// TIA Portal V20 export
FUNCTION_BLOCK "POS3_0_Antriebe"   // FB34, FBD
{ S7_Optimized_Access := 'TRUE' }
// stored: MemoryReserve 100, SetENOAutomatically false
   VAR
      "-1001T1_OM_PRM_Access_Instance" { S7_SetPoint := 'True'} : "OM_PRM_Access";
      "-1001T1_Oriental" { S7_SetPoint := 'True'} : "Oriental_AZD-KPN_Profinet";
      "-1002T2_OM_PRM_Access_Instance" { S7_SetPoint := 'True'} : "OM_PRM_Access";
      "-1002T2_Oriental_Drehachse" { S7_SetPoint := 'True'} : "Oriental_AZD-KPN_Profinet";
      Pos_Alt { S7_SetPoint := 'True'} : Real;
      Delta : Real;
   END_VAR
BEGIN

REGION Network 1 (SCL): -1001T1 Pos 3.0 Positionierachse Vorgaben Geschwindigkeit und Beschleunigung
   "POS3_0_Signal"."-1001T1 Oriental_Beschleunigung" := 50.0;
   "POS3_0_Signal"."-1001T1 Oriental_Speed" := 100.0;
END_REGION

REGION Network 2 (SCL): -1001T1 Pos 3.0 Positionierachse Achse stopp
   // Achse stopp
   IF "03_Betriebsart_DB"."Schutztüren OK" AND
       "DE_POS3_0_Endlage_Überlastzylinder" THEN
       "POS3_0_Signal"."-1001T1 Oriental_Steuerung".E_STOP := FALSE;
   ELSE
       "POS3_0_Signal"."-1001T1 Oriental_Steuerung".E_STOP := TRUE;
   END_IF;
END_REGION

REGION Network 3 (SCL): -1001T1 Pos 3.0 Positionierachse Position 0 Achse [Grundstellung]
   "POS3_0_Signal"."-1001T1 Oriental_Positionen".Operation_type[0] := 16#0001;
   "POS3_0_Signal"."-1001T1 Oriental_Positionen".Soll_Position[0] := 0.0;
   "POS3_0_Signal"."-1001T1 Oriental_Positionen".Geschwindigkeit[0] := 10.0;
   "POS3_0_Signal"."-1001T1 Oriental_Positionen".Start_Rampe[0] := "POS3_0_Signal"."-1001T1 Oriental_Beschleunigung"; // Start-Rampe %
   "POS3_0_Signal"."-1001T1 Oriental_Positionen".Stopp_Rampe[0] := "POS3_0_Signal"."-1001T1 Oriental_Beschleunigung"; // Stopp-Rampe %
   "POS3_0_Signal"."-1001T1 Oriental_Positionen".Arbeitsstrom[0] := 100;  // Arbeitsstrom in %
   "POS3_0_Signal"."-1001T1 Oriental_Positionen".Positioniertoleranz[0] := 0.02;
END_REGION

REGION Network 4 (SCL): -1001T1 Pos 3.0 Positionierachse Position 1 Achse [GS aus Verwaltung]
   "POS3_0_Signal"."-1001T1 Oriental_Positionen".Operation_type[1] := 16#0001;

   "POS3_0_Signal"."-1001T1 Oriental_Positionen".Start_Rampe[1] := "POS3_0_Signal"."-1001T1 Oriental_Beschleunigung"; // Start-Rampe %
   "POS3_0_Signal"."-1001T1 Oriental_Positionen".Stopp_Rampe[1] := "POS3_0_Signal"."-1001T1 Oriental_Beschleunigung"; // Stopp-Rampe %
   "POS3_0_Signal"."-1001T1 Oriental_Positionen".Arbeitsstrom[1] := 100;   // Arbeitsstrom in %
   "POS3_0_Signal"."-1001T1 Oriental_Positionen".Positioniertoleranz[1] := 0.02;
END_REGION

REGION Network 5 (SCL): -1001T1 Pos 3.0 Positionierachse Position 2 Achse [AS aus Verwaltung]
   "POS3_0_Signal"."-1001T1 Oriental_Positionen".Operation_type[2] := 16#0001;

   "POS3_0_Signal"."-1001T1 Oriental_Positionen".Start_Rampe[2] := "POS3_0_Signal"."-1001T1 Oriental_Beschleunigung"; // Start-Rampe %
   "POS3_0_Signal"."-1001T1 Oriental_Positionen".Stopp_Rampe[2] := "POS3_0_Signal"."-1001T1 Oriental_Beschleunigung"; // Stopp-Rampe %
   "POS3_0_Signal"."-1001T1 Oriental_Positionen".Arbeitsstrom[2] := 100;  // Arbeitsstrom in %
   "POS3_0_Signal"."-1001T1 Oriental_Positionen".Positioniertoleranz[2] := 0.02;
END_REGION

REGION Network 6 (SCL): -1001T1 Pos 3.0 Positionierachse Position 3 Achse
   "POS3_0_Signal"."-1001T1 Oriental_Positionen".Operation_type[3] := 16#0001;

   "POS3_0_Signal"."-1001T1 Oriental_Positionen".Start_Rampe[3] := "POS3_0_Signal"."-1001T1 Oriental_Beschleunigung" ; // Start-Rampe %
   "POS3_0_Signal"."-1001T1 Oriental_Positionen".Stopp_Rampe[3] := "POS3_0_Signal"."-1001T1 Oriental_Beschleunigung" ; // Stopp-Rampe %
   "POS3_0_Signal"."-1001T1 Oriental_Positionen".Arbeitsstrom[3] := 100; // Arbeitsstrom in %
   "POS3_0_Signal"."-1001T1 Oriental_Positionen".Positioniertoleranz[3] := 0.02;
END_REGION

REGION Network 7 (SCL): -1001T1 Pos 3.0 Positionierachse Position 4 Achse
   "POS3_0_Signal"."-1001T1 Oriental_Positionen".Operation_type[4] := 16#0001;

   "POS3_0_Signal"."-1001T1 Oriental_Positionen".Start_Rampe[4] := "POS3_0_Signal"."-1001T1 Oriental_Beschleunigung" ; // Start-Rampe %
   "POS3_0_Signal"."-1001T1 Oriental_Positionen".Stopp_Rampe[4] := "POS3_0_Signal"."-1001T1 Oriental_Beschleunigung" ; // Stopp-Rampe %
   "POS3_0_Signal"."-1001T1 Oriental_Positionen".Arbeitsstrom[4] := 100;  // Arbeitsstrom in %
   "POS3_0_Signal"."-1001T1 Oriental_Positionen".Positioniertoleranz[4] := 0.03;
END_REGION

REGION Network 8 (SCL): -1001T1 Pos 3.0 Positionierachse Position 5 Achse

   "POS3_0_Signal"."-1001T1 Oriental_Positionen".Operation_type[5] := 16#0001;

   "POS3_0_Signal"."-1001T1 Oriental_Positionen".Start_Rampe[5] := "POS3_0_Signal"."-1001T1 Oriental_Beschleunigung"; // Start-Rampe %
   "POS3_0_Signal"."-1001T1 Oriental_Positionen".Stopp_Rampe[5] := "POS3_0_Signal"."-1001T1 Oriental_Beschleunigung"; // Stopp-Rampe %
   "POS3_0_Signal"."-1001T1 Oriental_Positionen".Arbeitsstrom[5] := 100;  // Arbeitsstrom in %
   "POS3_0_Signal"."-1001T1 Oriental_Positionen".Positioniertoleranz[5] := 0.03;
END_REGION

REGION Network 9 (SCL): -1001T1 Pos 3.0 Positionierachse Grenzwerte
   "POS3_0_Signal"."-1001T1 Oriental_Positionen".A_Softw_ES_max_mm := 210.0;
   "POS3_0_Signal"."-1001T1 Oriental_Positionen".A_Softw_ES_min_mm := -0.5;
END_REGION

NETWORK
TITLE = -1001T1 Pos 3.0 Positionierachse E_ETO-CLR Quittieren nach "Sicherer Halt"
      A     "03_Betriebsart_DB"."NOT-HALT OK";
      A     "03_Betriebsart_DB"."Schutztüren OK";
      AN    "POS3_0_Signal"."-1001T1 Oriental_Steuerung"."A_DCMD-RDY";
      A     "FL_Clock_1Hz";
      =     "POS3_0_Signal"."-1001T1 Oriental_Steuerung"."E_ETO-CLR";


NETWORK
TITLE = -1001T1 Pos 3.0 Positionierachse Oriental Achse Parameter schreiben und lesen (wird nicht benötigt)
      CALL  #"-1001T1_OM_PRM_Access_Instance"
      ( Inputdata_RW_Drv2PLC  := "AZ_1001T1_Pos3_0__Prm_Status",
        ReadParameterID       := "POS3_0_Parameter_Data".RD_ParameterID,
        WriteParameterID      := "POS3_0_Parameter_Data".WR_ParameterID,
        WriteData             := "POS3_0_Parameter_Data".WR_ParameterData,
        "WR-REQ"              := ,
        Outputdata_RW_PLC2Drv := "AZ_1001T1_Pos3_0__Prm_Set",
        ReadParameterID_R     := ,
        WriteParameterID_R    := ,
        ReadData              := "POS3_0_Parameter_Data".RD_ParameterData,
        "WR-SET-ERR"          := ,
        "WR-IF-ERR"           := ,
        "WR-NV-ERR"           := ,
        "WR-EXE-ERR"          := ,
        "WR-ERR"              := ,
        "RD-ERR"              := ,
        "WR-END"              := ,
        "SYS-BSY"             := 
      );



REGION Network 12 (SCL): -1001T1 Pos 3.0 Positionierachse Oriental DDO_Type für E_Trig_Manuell
   // E_DDO_Type 16#0001 = absolut positionieren 16#0002 = relativ positionieren
   "POS3_0_Signal"."-1001T1 Oriental_Steuerung".E_DDO_Type := 16#0001;
END_REGION

NETWORK
TITLE = -1001T1 Pos 3.0 Positionierachse Oriental Achse Ansteuerung
      CALL  #"-1001T1_Oriental"
      ( Inputdata_FixedIO_Drv2PLC           := "AZ_1001T1_Pos3_0__Fixed_Out",
        MonitorData                         := "AZ_1001T1_Pos3_0__St_Monitor",
        E_DDO_Type                          := "POS3_0_Signal"."-1001T1 Oriental_Steuerung".E_DDO_Type,
        E_DDO_Pos                           := "POS3_0_Signal"."-1001T1 Oriental_Steuerung".E_DDO_Pos,
        E_DDO_Vel                           := "POS3_0_Signal"."-1001T1 Oriental_Steuerung".E_DDO_Vel,
        E_DDO_Acc                           := "POS3_0_Signal"."-1001T1 Oriental_Steuerung".E_DDO_Acc,
        E_DDO_Dec                           := "POS3_0_Signal"."-1001T1 Oriental_Steuerung".E_DDO_Dec,
        E_DDO_Crnt                          := "POS3_0_Signal"."-1001T1 Oriental_Steuerung".E_DDO_Crnt,
        E_DDO_Trans                         := "POS3_0_Signal"."-1001T1 Oriental_Steuerung".E_DDO_Trans,
        E_Schrittweite_Pos                  := "POS3_0_Signal"."-1001T1 Oriental_Steuerung".E_Schrittweite_pos,
        E_Schrittweite_Neg                  := "POS3_0_Signal"."-1001T1 Oriental_Steuerung".E_Schrittweite_neg,
        E_Schrittweite                      := "POS3_0_Signal"."-1001T1 Oriental_Steuerung".E_Schrittweite,
        E_R_Softw_ES_min_steps              := "POS3_0_Signal"."-1001T1 Oriental_Positionen".A_Softw_ES_min_mm,
        E_R_Softw_ES_max_steps              := "POS3_0_Signal"."-1001T1 Oriental_Positionen".A_Softw_ES_max_mm,
        E_Drehachse                         := FALSE,
        E_Getriebefaktor                    := 100.0,
        E_Maximalgeschwindigkeit_Hz         := 25000.0,
        "E_Maximal_Start_Stopp_Rampe_kHz/s" := 250000.0,
        E_SIMULATION_AKTIV                  := "03_Betriebsart_DB".Simulation_aktiv,
        E_RemoteIO                          := "AZ_1001T1_Pos3_0__Remote_Out",
        Outputdata_DDO                      := "AZ_1001T1_Pos3_0__DDO",
        Outputdata_FixedIO_PLC2Drv          := "AZ_1001T1_Pos3_0__Fixed_In",
        A_TRIG_R                            := "POS3_0_Signal"."-1001T1 Oriental_Steuerung".A_TRIG_R,
        "A_TRIG-MODE_R"                     := "POS3_0_Signal"."-1001T1 Oriental_Steuerung"."A_TRIG-MODE_R",
        "A_SET-ERR"                         := "POS3_0_Signal"."-1001T1 Oriental_Steuerung"."A_SET-ERR",
        "A_EXE-ERR"                         := "POS3_0_Signal"."-1001T1 Oriental_Steuerung"."A_EXE-ERR",
        "A_DCMD-FULL"                       := "POS3_0_Signal"."-1001T1 Oriental_Steuerung"."A_DCMD-FULL",
        A_STOP_R                            := "POS3_0_Signal"."-1001T1 Oriental_Steuerung".A_STOP_R,
        "A_ETO-MON"                         := "POS3_0_Signal"."-1001T1 Oriental_Steuerung"."A_ETO-MON",
        A_TLC                               := "POS3_0_Signal"."-1001T1 Oriental_Steuerung".A_TLC,
        "A_SEQ-BSY"                         := "POS3_0_Signal"."-1001T1 Oriental_Steuerung"."A_SEQ-BSY",
        A_MOVE                              := "POS3_0_Signal"."-1001T1 Oriental_Steuerung".A_MOVE,
        "A_IN-POS"                          := "POS3_0_Signal"."-1001T1 Oriental_Steuerung"."A_IN-POS",
        A_START_R                           := "POS3_0_Signal"."-1001T1 Oriental_Steuerung".A_START_R,
        "A_HOME-END"                        := "POS3_0_Signal"."-1001T1 Oriental_Steuerung"."A_HOME-END",
        A_READY                             := "POS3_0_Signal"."-1001T1 Oriental_Steuerung".A_READY,
        "A_DCMD-RDY"                        := "POS3_0_Signal"."-1001T1 Oriental_Steuerung"."A_DCMD-RDY",
        "A_ALM-A"                           := "POS3_0_Signal"."-1001T1 Oriental_Steuerung"."A_ALM-A",
        A_PresentAlarm                      := "POS3_0_Signal"."-1001T1 Oriental_Steuerung".A_PresentAlarm,
        A_FBposition                        := "POS3_0_Signal"."-1001T1 Oriental_Steuerung".A_FBposition,
        A_FBspeed                           := "POS3_0_Signal"."-1001T1 Oriental_Steuerung".A_FBspeed,
        A_CmdPosition                       := "POS3_0_Signal"."-1001T1 Oriental_Steuerung".A_CmdPosition,
        A_TorqueMonitor                     := "POS3_0_Signal"."-1001T1 Oriental_Steuerung".A_TorqueMonitor,
        A_CST_OpeCurrent                    := "POS3_0_Signal"."-1001T1 Oriental_Steuerung".A_CST_OpeCurrent,
        A_Information                       := "POS3_0_Signal"."-1001T1 Oriental_Steuerung".A_Information,
        A_StatusWord                        := "POS3_0_Signal"."-1001T1 Oriental_Steuerung".A_StatusWord,
        A_RemoteIO                          := "AZ_1001T1_Pos3_0__Remote_IN",
        E_A_UDT_Positionen                  := "POS3_0_Signal"."-1001T1 Oriental_Positionen",
        E_Not_Aus_OK                        := "03_Betriebsart_DB"."NOT-HALT OK",
        E_Tueren_OK                         := "03_Betriebsart_DB"."Schutztüren OK",
        "E_TRIG-MODE"                       := "POS3_0_Signal"."-1001T1 Oriental_Steuerung"."E_TRIG-MODE",
        "E_ETO-CLR"                         := "POS3_0_Signal"."-1001T1 Oriental_Steuerung"."E_ETO-CLR",
        "E_FW-JOG"                          := "POS3_0_Signal"."-1001T1 Oriental_Steuerung"."E_FW-JOG",
        "E_RV-JOG"                          := "POS3_0_Signal"."-1001T1 Oriental_Steuerung"."E_RV-JOG",
        E_START                             := "POS3_0_Signal"."-1001T1 Oriental_Steuerung".E_START,
        E_ZHOME                             := "POS3_0_Signal"."-1001T1 Oriental_Steuerung".E_ZHOME,
        E_STOP                              := "POS3_0_Signal"."-1001T1 Oriental_Steuerung".E_STOP,
        E_FREE                              := "POS3_0_Signal"."-1001T1 Oriental_Steuerung".E_FREE,
        "E_ALM-RST"                         := "03_Betriebsart_DB".ACK_Taste,
        E_TRIG_MANUELL                      := "POS3_0_Signal"."-1001T1 Oriental_Steuerung".E_Trig_Manuell,
        E_Home                              := "POS3_0_Signal"."-1001T1 Oriental_E_P-Preset"
      );

REGION Network 14 (SCL): -1001T1 Pos 3.0 "P-Preset" Reset
   IF "POS3_0_Signal"."-1001T1 Oriental_E_P-Preset" THEN
       "POS3_0_Signal"."-1001T1 Oriental_E_P-Preset" := False;
   END_IF;
END_REGION

REGION Network 16 (SCL): -1002T1 Pos 3.0 Drehachse Vorgaben Geschwindigkeit und Beschleunigung
   "POS3_0_Signal"."-1002T1_Oriental_Beschleunigung" := 40.0;
   "POS3_0_Signal"."-1002T1_Oriental_Speed" := 100.0;
END_REGION

REGION Network 17 (SCL): -1002T1 Pos 3.0 Drehachse Achse stopp
   // Achse stopp
   IF "03_Betriebsart_DB"."Schutztüren OK" THEN
       "POS3_0_Signal"."-1002T1 Oriental_Steuerung".E_STOP := FALSE;
   ELSE
       "POS3_0_Signal"."-1002T1 Oriental_Steuerung".E_STOP := TRUE;
   END_IF;
END_REGION

REGION Network 18 (SCL): -1002T1 Pos 3.0 Drehachse Position 0 [Grundstellung]
   "POS3_0_Signal"."-1002T1 Oriental_Positionen".Operation_type[0] := 16#0001;
   "POS3_0_Signal"."-1002T1 Oriental_Positionen".Soll_Position[0] := 0.0;
   "POS3_0_Signal"."-1002T1 Oriental_Positionen".Geschwindigkeit[0] := 10.0;
   "POS3_0_Signal"."-1002T1 Oriental_Positionen".Start_Rampe[0] := "POS3_0_Signal"."-1002T1_Oriental_Beschleunigung"; // Start-Rampe %
   "POS3_0_Signal"."-1002T1 Oriental_Positionen".Stopp_Rampe[0] := "POS3_0_Signal"."-1002T1_Oriental_Beschleunigung"; // Stopp-Rampe %
   "POS3_0_Signal"."-1002T1 Oriental_Positionen".Arbeitsstrom[0] := 100;  // Arbeitsstrom in %
   "POS3_0_Signal"."-1002T1 Oriental_Positionen".Positioniertoleranz[0] := 0.001;
END_REGION

REGION Network 19 (SCL): -1002T1 Pos 3.0 Drehachse Position 1 [0.0 ° Absolut positionieren]
   "POS3_0_Signal"."-1002T1 Oriental_Positionen".Operation_type[1] := 16#0001;
   "POS3_0_Signal"."-1002T1 Oriental_Positionen".Soll_Position[1] := 0.0;
   "POS3_0_Signal"."-1002T1 Oriental_Positionen".Geschwindigkeit[1] := 10.0;
   "POS3_0_Signal"."-1002T1 Oriental_Positionen".Start_Rampe[1] := "POS3_0_Signal"."-1002T1_Oriental_Beschleunigung"; // Start-Rampe %
   "POS3_0_Signal"."-1002T1 Oriental_Positionen".Stopp_Rampe[1] := "POS3_0_Signal"."-1002T1_Oriental_Beschleunigung"; // Stopp-Rampe %
   "POS3_0_Signal"."-1002T1 Oriental_Positionen".Arbeitsstrom[1] := 100;   // Arbeitsstrom in %
   "POS3_0_Signal"."-1002T1 Oriental_Positionen".Positioniertoleranz[1] := 0.001;
END_REGION

REGION Network 20 (SCL): -1002T1 Pos 3.0 Drehachse Position 2 [AS1 aus Verwaltung]
   "POS3_0_Signal"."-1002T1 Oriental_Positionen".Operation_type[2] := 16#0002;

   "POS3_0_Signal"."-1002T1 Oriental_Positionen".Start_Rampe[2] := "POS3_0_Signal"."-1002T1_Oriental_Beschleunigung"; // Start-Rampe %
   "POS3_0_Signal"."-1002T1 Oriental_Positionen".Stopp_Rampe[2] := "POS3_0_Signal"."-1002T1_Oriental_Beschleunigung"; // Stopp-Rampe %
   "POS3_0_Signal"."-1002T1 Oriental_Positionen".Arbeitsstrom[2] := REAL_TO_DINT ("Verwaltung_Teiledaten"."Drehantrieb Motorstrombegrenzung");  // Arbeitsstrom in %
   "POS3_0_Signal"."-1002T1 Oriental_Positionen".Positioniertoleranz[2] := 0.001;
END_REGION

REGION Network 21 (SCL): -1002T1 Pos 3.0 Drehachse Position 3 [GS aus Verwaltung]
   "POS3_0_Signal"."-1002T1 Oriental_Positionen".Operation_type[3] := 16#0002;

   "POS3_0_Signal"."-1002T1 Oriental_Positionen".Start_Rampe[3] := "POS3_0_Signal"."-1002T1_Oriental_Beschleunigung"; // Start-Rampe %
   "POS3_0_Signal"."-1002T1 Oriental_Positionen".Stopp_Rampe[3] := "POS3_0_Signal"."-1002T1_Oriental_Beschleunigung"; // Stopp-Rampe %
   "POS3_0_Signal"."-1002T1 Oriental_Positionen".Arbeitsstrom[3] := REAL_TO_DINT ("Verwaltung_Teiledaten"."Drehantrieb Motorstrombegrenzung");  // Arbeitsstrom in %
   "POS3_0_Signal"."-1002T1 Oriental_Positionen".Positioniertoleranz[3] := 0.001;
END_REGION

REGION Network 22 (SCL): -1002T1 Pos 3.0 Drehachse Position 4
   "POS3_0_Signal"."-1002T1 Oriental_Positionen".Operation_type[4] := 16#0001;

   "POS3_0_Signal"."-1002T1 Oriental_Positionen".Start_Rampe[4] := "POS3_0_Signal"."-1002T1_Oriental_Beschleunigung"; // Start-Rampe %
   "POS3_0_Signal"."-1002T1 Oriental_Positionen".Stopp_Rampe[4] := "POS3_0_Signal"."-1002T1_Oriental_Beschleunigung"; // Stopp-Rampe %
   "POS3_0_Signal"."-1002T1 Oriental_Positionen".Arbeitsstrom[4] := 100;  // Arbeitsstrom in %
   "POS3_0_Signal"."-1002T1 Oriental_Positionen".Positioniertoleranz[4] := 0.01;
END_REGION

REGION Network 23 (SCL): -1002T1 Pos 3.0 Drehachse Position 5
   "POS3_0_Signal"."-1002T1 Oriental_Positionen".Operation_type[5] := 16#0001;

   "POS3_0_Signal"."-1002T1 Oriental_Positionen".Start_Rampe[5] := "POS3_0_Signal"."-1002T1_Oriental_Beschleunigung"; // Start-Rampe %
   "POS3_0_Signal"."-1002T1 Oriental_Positionen".Stopp_Rampe[5] := "POS3_0_Signal"."-1002T1_Oriental_Beschleunigung"; // Stopp-Rampe %
   "POS3_0_Signal"."-1002T1 Oriental_Positionen".Arbeitsstrom[5] := 100;  // Arbeitsstrom in %
   "POS3_0_Signal"."-1002T1 Oriental_Positionen".Positioniertoleranz[5] := 0.01;
END_REGION

REGION Network 24 (SCL): -1002T1 Pos 3.0 Drehachse Grenzwerte
   "POS3_0_Signal"."-1002T1 Oriental_Positionen".A_Softw_ES_max_mm := 10000.5;
   "POS3_0_Signal"."-1002T1 Oriental_Positionen".A_Softw_ES_min_mm := -10000.5;
END_REGION

NETWORK
TITLE = -1002T1 Pos 3.0 Drehachse E_ETO-CLR Quittieren nach "Sicherer Halt"
      A     "03_Betriebsart_DB"."NOT-HALT OK";
      A     "03_Betriebsart_DB"."Schutztüren OK";
      AN    "POS3_0_Signal"."-1002T1 Oriental_Steuerung"."A_DCMD-RDY";
      A     "FL_Clock_1Hz";
      =     "POS3_0_Signal"."-1002T1 Oriental_Steuerung"."E_ETO-CLR";


NETWORK
TITLE = -1002T1 Pos 3.0 Drehachse Oriental Achse Parameter schreiben und lesen (wird nicht benötigt)
      CALL  #"-1002T2_OM_PRM_Access_Instance"
      ( Inputdata_RW_Drv2PLC  := "AZ_1002T1_Pos3_0_Drehachse__Prm_Status",
        ReadParameterID       := "POS3_0_Parameter_Data_Drehachse".RD_ParameterID,
        WriteParameterID      := "POS3_0_Parameter_Data_Drehachse".WR_ParameterID,
        WriteData             := "POS3_0_Parameter_Data_Drehachse".WR_ParameterData,
        "WR-REQ"              := ,
        Outputdata_RW_PLC2Drv := "AZ_1002T1_Pos3_0_Drehachse__Prm_Set",
        ReadParameterID_R     := ,
        WriteParameterID_R    := ,
        ReadData              := "POS3_0_Parameter_Data_Drehachse".RD_ParameterData,
        "WR-SET-ERR"          := ,
        "WR-IF-ERR"           := ,
        "WR-NV-ERR"           := ,
        "WR-EXE-ERR"          := ,
        "WR-ERR"              := ,
        "RD-ERR"              := ,
        "WR-END"              := ,
        "SYS-BSY"             := 
      );



REGION Network 27 (SCL): -1002T1 Pos 3.0 Drehachse DDO_Type für E_Trig_Manuell
   // E_DDO_Type 16#0001 = absolut positionieren 16#0002 = relativ positionieren
   "POS3_0_Signal"."-1002T1 Oriental_Steuerung".E_DDO_Type := 16#0002;
END_REGION

NETWORK
TITLE = -1002T1 Pos 3.0 Drehachse Oriental Achse Ansteuerung
      CALL  #"-1002T2_Oriental_Drehachse"
      ( Inputdata_FixedIO_Drv2PLC           := "AZ_1002T1_Pos3_0_Drehachse__Fixed_Out",
        MonitorData                         := "AZ_1002T1_Pos3_0_Drehachse__St_Monitor",
        E_DDO_Type                          := "POS3_0_Signal"."-1002T1 Oriental_Steuerung".E_DDO_Type,
        E_DDO_Pos                           := "POS3_0_Signal"."-1002T1 Oriental_Steuerung".E_DDO_Pos,
        E_DDO_Vel                           := "POS3_0_Signal"."-1002T1 Oriental_Steuerung".E_DDO_Vel,
        E_DDO_Acc                           := "POS3_0_Signal"."-1002T1 Oriental_Steuerung".E_DDO_Acc,
        E_DDO_Dec                           := "POS3_0_Signal"."-1002T1 Oriental_Steuerung".E_DDO_Dec,
        E_DDO_Crnt                          := "POS3_0_Signal"."-1002T1 Oriental_Steuerung".E_DDO_Crnt,
        E_DDO_Trans                         := "POS3_0_Signal"."-1002T1 Oriental_Steuerung".E_DDO_Trans,
        E_Schrittweite_Pos                  := "POS3_0_Signal"."-1002T1 Oriental_Steuerung".E_Schrittweite_pos,
        E_Schrittweite_Neg                  := "POS3_0_Signal"."-1002T1 Oriental_Steuerung".E_Schrittweite_neg,
        E_Schrittweite                      := "POS3_0_Signal"."-1002T1 Oriental_Steuerung".E_Schrittweite,
        E_R_Softw_ES_min_steps              := "POS3_0_Signal"."-1002T1 Oriental_Positionen".A_Softw_ES_min_mm,
        E_R_Softw_ES_max_steps              := "POS3_0_Signal"."-1002T1 Oriental_Positionen".A_Softw_ES_max_mm,
        E_Drehachse                         := TRUE,
        E_Getriebefaktor                    := 18.0,
        E_Maximalgeschwindigkeit_Hz         := 30000.0,
        "E_Maximal_Start_Stopp_Rampe_kHz/s" := 990000.0,
        E_SIMULATION_AKTIV                  := "03_Betriebsart_DB".Simulation_aktiv,
        E_RemoteIO                          := "AZ_1002T1_Pos3_0_Drehachse__Remote_Out",
        Outputdata_DDO                      := "AZ_1002T1_Pos3_0_Drehachse__DDO",
        Outputdata_FixedIO_PLC2Drv          := "AZ_1002T1_Pos3_0_Drehachse__Fixed_In",
        A_TRIG_R                            := "POS3_0_Signal"."-1002T1 Oriental_Steuerung".A_TRIG_R,
        "A_TRIG-MODE_R"                     := "POS3_0_Signal"."-1002T1 Oriental_Steuerung"."A_TRIG-MODE_R",
        "A_SET-ERR"                         := "POS3_0_Signal"."-1002T1 Oriental_Steuerung"."A_SET-ERR",
        "A_EXE-ERR"                         := "POS3_0_Signal"."-1002T1 Oriental_Steuerung"."A_EXE-ERR",
        "A_DCMD-FULL"                       := "POS3_0_Signal"."-1002T1 Oriental_Steuerung"."A_DCMD-FULL",
        A_STOP_R                            := "POS3_0_Signal"."-1002T1 Oriental_Steuerung".A_STOP_R,
        "A_ETO-MON"                         := "POS3_0_Signal"."-1002T1 Oriental_Steuerung"."A_ETO-MON",
        A_TLC                               := "POS3_0_Signal"."-1002T1 Oriental_Steuerung".A_TLC,
        "A_SEQ-BSY"                         := "POS3_0_Signal"."-1002T1 Oriental_Steuerung"."A_SEQ-BSY",
        A_MOVE                              := "POS3_0_Signal"."-1002T1 Oriental_Steuerung".A_MOVE,
        "A_IN-POS"                          := "POS3_0_Signal"."-1002T1 Oriental_Steuerung"."A_IN-POS",
        A_START_R                           := "POS3_0_Signal"."-1002T1 Oriental_Steuerung".A_START_R,
        "A_HOME-END"                        := "POS3_0_Signal"."-1002T1 Oriental_Steuerung"."A_HOME-END",
        A_READY                             := "POS3_0_Signal"."-1002T1 Oriental_Steuerung".A_READY,
        "A_DCMD-RDY"                        := "POS3_0_Signal"."-1002T1 Oriental_Steuerung"."A_DCMD-RDY",
        "A_ALM-A"                           := "POS3_0_Signal"."-1002T1 Oriental_Steuerung"."A_ALM-A",
        A_PresentAlarm                      := "POS3_0_Signal"."-1002T1 Oriental_Steuerung".A_PresentAlarm,
        A_FBposition                        := "POS3_0_Signal"."-1002T1 Oriental_Steuerung".A_FBposition,
        A_FBspeed                           := "POS3_0_Signal"."-1002T1 Oriental_Steuerung".A_FBspeed,
        A_CmdPosition                       := "POS3_0_Signal"."-1002T1 Oriental_Steuerung".A_CmdPosition,
        A_TorqueMonitor                     := "POS3_0_Signal"."-1002T1 Oriental_Steuerung".A_TorqueMonitor,
        A_CST_OpeCurrent                    := "POS3_0_Signal"."-1002T1 Oriental_Steuerung".A_CST_OpeCurrent,
        A_Information                       := "POS3_0_Signal"."-1002T1 Oriental_Steuerung".A_Information,
        A_StatusWord                        := "POS3_0_Signal"."-1002T1 Oriental_Steuerung".A_StatusWord,
        A_RemoteIO                          := "AZ_1002T1_Pos3_0_Drehachse__Remote_IN",
        E_A_UDT_Positionen                  := "POS3_0_Signal"."-1002T1 Oriental_Positionen",
        E_Not_Aus_OK                        := "03_Betriebsart_DB"."NOT-HALT OK",
        E_Tueren_OK                         := "03_Betriebsart_DB"."Schutztüren OK",
        "E_TRIG-MODE"                       := "POS3_0_Signal"."-1002T1 Oriental_Steuerung"."E_TRIG-MODE",
        "E_ETO-CLR"                         := "POS3_0_Signal"."-1002T1 Oriental_Steuerung"."E_ETO-CLR",
        "E_FW-JOG"                          := "POS3_0_Signal"."-1002T1 Oriental_Steuerung"."E_FW-JOG",
        "E_RV-JOG"                          := "POS3_0_Signal"."-1002T1 Oriental_Steuerung"."E_RV-JOG",
        E_START                             := "POS3_0_Signal"."-1002T1 Oriental_Steuerung".E_START,
        E_ZHOME                             := "POS3_0_Signal"."-1002T1 Oriental_Steuerung".E_ZHOME,
        E_STOP                              := "POS3_0_Signal"."-1002T1 Oriental_Steuerung".E_STOP,
        E_FREE                              := "POS3_0_Signal"."-1002T1 Oriental_Steuerung".E_FREE,
        "E_ALM-RST"                         := "03_Betriebsart_DB".ACK_Taste,
        E_TRIG_MANUELL                      := "POS3_0_Signal"."-1002T1 Oriental_Steuerung".E_Trig_Manuell,
        E_Home                              := "POS3_0_Signal"."-1002T1 Oriental_E_P-Preset"
      );

REGION Network 29 (SCL): -1002T1 Pos 3.0 Drehachse "P-Preset" Reset
   IF "POS3_0_Signal"."-1002T1 Oriental_E_P-Preset" THEN
       "POS3_0_Signal"."-1002T1 Oriental_E_P-Preset" := False;
       "POS3_0_Signal"."-1002T1 Oriental_Umdrehungszähler" := 0.0;
   END_IF;
END_REGION

REGION Network 30 (SCL): -1002T1 Pos 3.0 Drehachse Berechnung der Umdrehungen ab dem Nullpunkt
   // Positionsdifferenz berechnen
   #Delta := "POS3_0_Signal"."-1002T1 Oriental_Steuerung".A_FBposition - #Pos_Alt;

   //Überlauf erkennen 
   IF #Delta < -180.0 THEN
       // Vorwärts über 360° gelaufen (z.B. 359 -> 1)
       "POS3_0_Signal"."-1002T1 Oriental_Umdrehungszähler" :=
       "POS3_0_Signal"."-1002T1 Oriental_Umdrehungszähler" + 1.0;

   ELSIF #Delta > 180.0 THEN
       // Rückwärts über 0° gelaufen (z.B. 1 -> 359)    
       "POS3_0_Signal"."-1002T1 Oriental_Umdrehungszähler" :=
       "POS3_0_Signal"."-1002T1 Oriental_Umdrehungszähler" - 1.0;
   END_IF;

   // Aktuellen Wert für nächsten Zyklus speichern
   #Pos_Alt := "POS3_0_Signal"."-1002T1 Oriental_Steuerung".A_FBposition;


   "POS3_0_Signal"."-1002T1 Oriental_Absolute_Position" :=    "POS3_0_Signal"."-1002T1 Oriental_Umdrehungszähler" * 360.0 +
   "POS3_0_Signal"."-1002T1 Oriental_Steuerung".A_FBposition;
END_REGION

REGION Network 31 (SCL): -1002T1 Pos 3.0 Drehachse Kraft überschritten
   IF "POS3_0_Signal"."-1002T1 Oriental_Steuerung".A_TorqueMonitor >=
      "POS3_0_Signal"."-1002T1 Oriental_Steuerung".A_CST_OpeCurrent   THEN
       "POS3_0_Signal".Drehachse_Kraft_überschritten := true;
   ELSE
       "POS3_0_Signal".Drehachse_Kraft_überschritten := false;
   END_IF;
END_REGION
END_FUNCTION_BLOCK
